(* IEC 61131-3 sources: STAR-PLC-Agent/results/raw/four_group_20261114/star_deepseek_v4/SELF002/formal/attempt_0001, 1 file *)

(* ---- candidate.st ---- *)
FUNCTION_BLOCK FB_Task
VAR_INPUT
    ForwardButton : BOOL;
    ReverseButton : BOOL;
    Stop : BOOL;
END_VAR
VAR_OUTPUT
    Forward : BOOL := FALSE;
    Reverse : BOOL := FALSE;
END_VAR
VAR
    previous_direction : INT := 0;
    desired_direction : INT := 0;
END_VAR

desired_direction := 0;
IF Stop OR (ForwardButton = ReverseButton) THEN
    desired_direction := 0;
ELSIF ForwardButton THEN
    desired_direction := 1;
ELSIF ReverseButton THEN
    desired_direction := -1;
END_IF;

IF (desired_direction <> 0) AND (previous_direction <> 0) AND (desired_direction <> previous_direction) THEN
    Forward := FALSE;
    Reverse := FALSE;
    previous_direction := 0;
ELSE
    Forward := (desired_direction = 1);
    Reverse := (desired_direction = -1);
    previous_direction := desired_direction;
END_IF;
END_FUNCTION_BLOCK
